// TIA Portal project "000_empty" (V21)

(* hardware
DEVICE "PLC_1"  S7-1500 station
   slot 0: "Rail_0"  Rack  6ES7 590-1***0-0AA0
   slot 1: "PLC_1"  CPU 1513-1 PN  6ES7 513-1AL02-0AB0  V2.9
      slot 3: "CPU display_1"  6ES7591-1AA00-0AA0
      slot 32768: "PROFINET interface_1"  X1
         slot 32769: "Port_1"  X1 P1
         slot 32770: "Port_2"  X1 P2
      slot 34817: "Virtual CP interface port_1"  Virtual CP interface port  Virtual CP interface port
*)

// ===== PLC "PLC_1"  CPU 1513-1 PN =====

VAR_GLOBAL   // PLC tag table "Default tag table"
   "tBool" AT %M0.0 : Bool;
   "tBool2" AT %M0.1 : Bool;
   "tInt" AT %MW2 : Int;
   "tDInt" AT %MD4 : DInt;
   "tReal" AT %MD8 : Real;
   "tWord" AT %MW12 : Word;
   "tByte" AT %MB14 : Byte;
   "tDWord" AT %MD16 : DWord;
   "tTime" AT %MD20 : Time;
   "tIn" AT %I0.0 : Bool;
   "tOut" AT %Q0.0 : Bool;
   "tUInt" AT %MW24 : UInt;
   "tLReal" AT %MD26 : LReal;
   "Tag_1" AT %MW100 : Word;
   "Tag_2" AT %M10.3 : Bool;
   "Tag_3" AT %Q1.0 : Bool;
   "Tag_4" AT %I1.0 : Bool;
   "Tag_5" AT %MD104 : DWord;
   "Tag_6" AT %MB110 : Byte;
   "Tag_7" AT %IW0 : Word;
   "Tag_8" AT %QW0 : Word;
END_VAR

VAR_GLOBAL CONSTANT   // PLC tag table "Default tag table"
   "MAX_COUNT" : Int := 100;
   "GAIN" : Real := 2.5;
   "TXT" : String := 'abc';
END_VAR

TYPE "UDT_Motor"
   STRUCT
      Running : Bool;   // Motor on
      Speed : Real := 1500.0;   // Speed setpoint
      Count : Int := 7;
   END_STRUCT;
END_TYPE

DATA_BLOCK "DB_Global"   // DB1
{ S7_Optimized_Access := 'TRUE' }
   VAR
      xBool : Bool := TRUE;   // Bool comment
      iInt : Int := 42;
      rReal : Real := 3.5;   // Real comment
      aInt : Array[0..3] of Int;
      sData : Struct
         "a" : Bool;
         "b" : DInt := -5;
      END_STRUCT;
   END_VAR
BEGIN
   aInt[1] := 11;
END_DATA_BLOCK

DATA_BLOCK "FB_Empty_DB"   // DB2
{ S7_Optimized_Access := 'TRUE' }
VERSION : 0.1
// stored: InstanceOfName FB_Empty
"FB_Empty"
BEGIN
END_DATA_BLOCK

DATA_BLOCK "DB_Motor"   // DB4
{ S7_Optimized_Access := 'TRUE' }
   VAR
      motor : "UDT_Motor";
   END_VAR
BEGIN
   motor.Speed := 750.0;
END_DATA_BLOCK

DATA_BLOCK "FB_Iface_DB"   // DB5
{ S7_Optimized_Access := 'TRUE' }
VERSION : 0.1
// stored: InstanceOfName FB_Iface
"FB_Iface"
BEGIN
   stInt := 99;
   stBool := TRUE;
END_DATA_BLOCK

DATA_BLOCK "DB_Std"   // DB6
{ S7_Optimized_Access := 'FALSE' }
   VAR
      x : Bool;
      i : Int;
      d : DInt;
      r : Real;
      "by" : Byte;
   END_VAR
BEGIN
END_DATA_BLOCK

// folder: BlockGroup_1

DATA_BLOCK "DB_InGroup"   // DB3
{ S7_Optimized_Access := 'TRUE' }
   VAR
      wWord : Word := 16#00FF;
   END_VAR
BEGIN
END_DATA_BLOCK

// folder: (top level)

DATA_BLOCK "TO_Speed_5_0"   // DB8, Motion_DB
{ S7_Optimized_Access := 'TRUE' }
AUTHOR : SIMATIC
FAMILY : MC_1500
VERSION : 5.0
// stored: InstanceOfName TO_SpeedAxis
"TO_SpeedAxis"
BEGIN
END_DATA_BLOCK

DATA_BLOCK "TO_Posit_6_0"   // DB10, Motion_DB
{ S7_Optimized_Access := 'TRUE' }
AUTHOR : SIMATIC
FAMILY : MC_1500
VERSION : 6.0
// stored: InstanceOfName TO_PositioningAxis
"TO_PositioningAxis"
BEGIN
END_DATA_BLOCK

DATA_BLOCK "TO_Exter_6_0"   // DB13, Motion_DB
{ S7_Optimized_Access := 'TRUE' }
AUTHOR : SIMATIC
FAMILY : MC_1500
VERSION : 6.0
// stored: InstanceOfName TO_ExternalEncoder
"TO_ExternalEncoder"
BEGIN
END_DATA_BLOCK

DATA_BLOCK "SpeedAx_6_0"   // DB14, Motion_DB
{ S7_Optimized_Access := 'TRUE' }
AUTHOR : SIMATIC
FAMILY : MC_1500
VERSION : 6.0
// stored: InstanceOfName TO_SpeedAxis
"TO_SpeedAxis"
BEGIN
END_DATA_BLOCK

FUNCTION_BLOCK "FB_Empty"   // FB1, SCL
{ S7_Optimized_Access := 'TRUE' }
VERSION : 0.1
BEGIN
END_FUNCTION_BLOCK

FUNCTION_BLOCK "FB_Iface"   // FB2, SCL
{ S7_Optimized_Access := 'TRUE' }
VERSION : 0.1
   VAR_INPUT
      iBool : Bool;   // Input bool
      iInt : Int;   // Input int
      iReal : Real;   // Input real
      iArr : Array[0..3] of Int;   // Input array
      iMotor : "UDT_Motor";   // Input UDT
   END_VAR
   VAR_OUTPUT
      oBool : Bool;   // Output bool
      oInt : Int;   // Output int
   END_VAR
   VAR_IN_OUT
      ioReal : Real;   // InOut real
   END_VAR
   VAR
      stInt : Int := 42;   // Static int
      stBool : Bool;   // Static bool comment
   END_VAR
   VAR_TEMP
      tInt : Int;   // Temp int
   END_VAR
   VAR CONSTANT
      cInt : Int := 7;   // Constant int
   END_VAR
BEGIN
   #tInt := #iInt + #cInt;
           #oInt := #tInt;
           #oBool := #iBool;
           #ioReal := #ioReal + #iReal;
END_FUNCTION_BLOCK

FUNCTION_BLOCK "FB_SclCalls"   // FB3, SCL
{ S7_Optimized_Access := 'TRUE' }
VERSION : 0.1
   VAR_INPUT
      start : Bool;
      pt : Time;
   END_VAR
   VAR_OUTPUT
      q : Bool;
      cnt : Int;
   END_VAR
   VAR
      tonInst : TON_TIME;
      tofInst : TOF_TIME;
      tpInst : TP_TIME;
      ctuInst : CTU_INT;
      trig : R_TRIG;
      ftrig : F_TRIG;
      "counter" : Int;
      ifc : "FB_Iface";
   END_VAR
   VAR_TEMP
      r : Real;
      "b" : Bool;
      res : Int;
      tot : Int;
   END_VAR
BEGIN
   #tonInst(IN := #start, PT := #pt);
   #q := #tonInst.Q;
   #tofInst(IN := #start, PT := T#2s);
   #tpInst(IN := #start, PT := #pt, Q => #b);
   #ctuInst(CU := #start, R := FALSE, PV := 10);
   #cnt := #ctuInst.CV;
   #trig(CLK := #start);
   IF #trig.Q THEN
       #counter := 0;
   END_IF;
   #ftrig(CLK := #start);
   #b := #ftrig.Q;
   #ifc(iBool := TRUE, iInt := 2, iReal := 1.0, ioReal := #r);
   #cnt := #ifc.oInt;
   "FB_Iface_DB"(iBool := #start, iInt := #cnt, iReal := #r, ioReal := #r, oInt => #cnt);
   "FC_SclOps"();
   #res := "FC_SclCtl"(n := 5, flag := TRUE, total => #tot);
   #res := "FC_SclCtl"(n := #res, flag := #b, total => #tot);
END_FUNCTION_BLOCK

FUNCTION_BLOCK "FB_SclLocal"   // FB4, SCL
{ S7_Optimized_Access := 'TRUE' }
VERSION : 0.1
   VAR_INPUT
      start : Bool;
   END_VAR
   VAR_IN_OUT
      io : Int;
   END_VAR
   VAR
      "counter" : Int;
      arr : Array[0..9] of Int;
      arr2 : Array[1..3, 1..4] of Real;
      mot : "UDT_Motor";
      st : Struct
         "a" : Int;
         "b" : Real;
         c : Array[0..2] of Bool;
      END_STRUCT;
   END_VAR
   VAR_TEMP
      i : Int;
   END_VAR
BEGIN
   #arr[0] := 1;
   #arr[#i] := #arr[#i + 1] + #io;
   #arr2[2, 3] := 1.5;
   #st.a := 10;
   #st.b := #st.a;
   #st.c[1] := TRUE;
   #mot.Speed := 100.0;
   #mot.Running := #st.c[0];
   #counter += 1;
   #io := #counter;
END_FUNCTION_BLOCK

FUNCTION_BLOCK "FB_LadTech"   // FB5, LAD
{ S7_Optimized_Access := 'TRUE' }
   VAR_INPUT
      sp : Real;
      pv : Real;
   END_VAR
   VAR_OUTPUT
      outv : Real;
      err : Bool;
   END_VAR
BEGIN

REGION Network 1: PID call
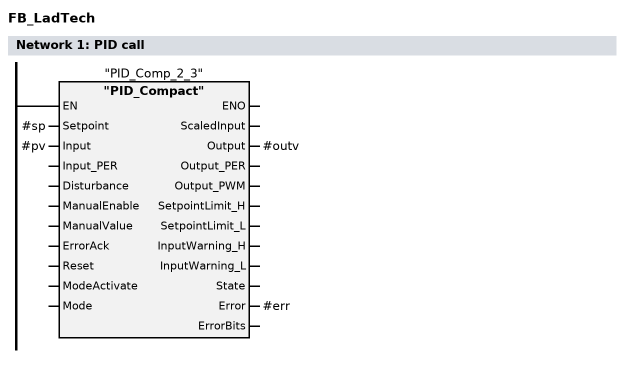
   RUNG wire#powerrail
      "PID_Comp_2_3"(Setpoint := #sp, Input := #pv, Output => #outv, Error => #err, Input_PER :=, Disturbance :=, ManualEnable :=, ManualValue :=, ErrorAck :=, Reset :=, ModeActivate :=, ScaledInput =>, Output_PER =>, Output_PWM =>, SetpointLimit_H =>, SetpointLimit_L =>, InputWarning_H =>, InputWarning_L =>, State =>, ErrorBits =>, Mode :=)
   END_RUNG
   // the same network as SCL:
   "PID_Comp_2_3"(Setpoint := #sp, Input := #pv, Output => #outv, Error => #err);   // "PID_Compact"
END_REGION
END_FUNCTION_BLOCK

FUNCTION_BLOCK "FB_FbdTech"   // FB6, FBD
{ S7_Optimized_Access := 'TRUE' }
   VAR_INPUT
      sp : Real;
      pv : Real;
   END_VAR
   VAR_OUTPUT
      outv : Real;
      err : Bool;
   END_VAR
BEGIN

REGION Network 1: PID call
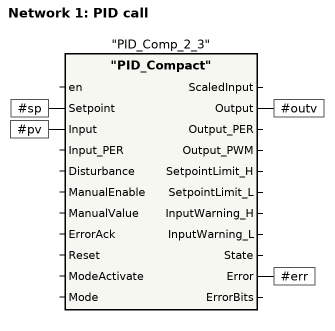
   "PID_Comp_2_3"(Setpoint := #sp, Input := #pv, Output => #outv, Error => #err);   // "PID_Compact"
END_REGION
END_FUNCTION_BLOCK

FUNCTION_BLOCK "FB_SclTech"   // FB7, SCL
{ S7_Optimized_Access := 'TRUE' }
   VAR_INPUT
      sp : Real;
      pv : Real;
   END_VAR
   VAR_OUTPUT
      outv : Real;
      err : Bool;
   END_VAR
BEGIN
// PID call
   "PID_Comp_2_3"(Setpoint := #sp, Input := #pv, Output => #outv, Error => #err);
END_FUNCTION_BLOCK

FUNCTION "FC_SclOps" : Void   // FC1, SCL
{ S7_Optimized_Access := 'TRUE' }
VERSION : 0.1
   VAR_TEMP
      b1 : Bool;
      b2 : Bool;
      b3 : Bool;
      i1 : Int;
      i2 : Int;
      i3 : Int;
      d1 : DInt;
      r1 : Real;
      r2 : Real;
      l1 : LReal;
      w1 : Word;
      w2 : Word;
      dw1 : DWord;
      by1 : Byte;
      u1 : UInt;
   END_VAR
BEGIN
   // arithmetic
           #i1 := 1 + 2 - 3 * 4;
           #i2 := #i1 / 2;
           #i3 := #i1 MOD 3;
           #r1 := #r2 ** 2.0;
           #i1 := -#i2;
           #i1 := +#i2;
           #i1 := (#i2 + #i3) * (#i2 - #i3);
           #d1 := #i1 * #i2;
           #r1 := #r2 / 3.0;
           #u1 := 5;
           // logic
           #b1 := NOT #b2;
           #b1 := #b2 AND #b3;
           #b1 := #b2 OR #b3;
           #b1 := #b2 XOR #b3;
           #b1 := #b2 & #b3;
           #b1 := (#b2 AND #b3) OR NOT (#b2 XOR #b3);
           #w1 := #w1 AND #w2;
           #w1 := #w1 OR #w2;
           #w1 := #w1 XOR #w2;
           #w1 := NOT #w2;
           // comparison
           #b1 := #i1 = #i2;
           #b1 := #i1 <> #i2;
           #b1 := #i1 < #i2;
           #b1 := #i1 <= #i2;
           #b1 := #i1 > #i2;
           #b1 := #i1 >= #i2;
           #b1 := #r1 > 1.5 AND #r2 <= 2.5;
           // compound assignment
           #i1 += 1;
           #i1 -= 1;
           #i1 *= 2;
           #i1 /= 2;
           // mixed types
           #l1 := #r1 + #d1;
           #r1 := #i1;
           #by1 := 16#FF;
           #dw1 := 16#DEADBEEF;
           #w1 := 2#1010_1010;
           #i1 := 8#17;
           #r1 := 1.0E3;
           #r2 := 2.5e-3;
           #l1 := 3.141592653589793;
END_FUNCTION

FUNCTION "FC_SclCtl" : Int   // FC2, SCL
{ S7_Optimized_Access := 'TRUE' }
VERSION : 0.1
   VAR_INPUT
      n : Int;
      flag : Bool;
   END_VAR
   VAR_OUTPUT
      total : Int;
   END_VAR
   VAR_TEMP
      i : Int;
      j : Int;
      x : Int;
      "b" : Bool;
   END_VAR
BEGIN
   (* block comment
      over two lines *)
   #total := 0;
   // IF forms
   IF #flag THEN
       #total := 1;
   END_IF;
   IF #n > 5 THEN
       #total := 2;
   ELSE
       #total := 3;
   END_IF;
   IF #n > 10 THEN
       #total := 4;
   ELSIF #n > 5 THEN
       #total := 5;
   ELSIF #n > 0 THEN
       #total := 6;
   ELSE
       #total := 7;
   END_IF;
   // CASE
   CASE #n OF
       0:
           #total := 10;
       1, 2:
           #total := 11;
       3..5:
           #total := 12;
       6, 8..9:
           #total := 13;
   ELSE
       #total := 14;
   END_CASE;
   CASE #x OF
       1:
           ;
   END_CASE;
   // FOR with BY, EXIT, CONTINUE
   FOR #i := 0 TO 10 DO
       #total += #i;
   END_FOR;
   FOR #i := 10 TO 0 BY -2 DO
       IF #i = 4 THEN
           CONTINUE;
       END_IF;
       IF #i = 2 THEN
           EXIT;
       END_IF;
       #total += #i;
   END_FOR;
   // nested loops
   FOR #i := 1 TO 3 DO
       FOR #j := 1 TO 3 DO
           #total := #total + #i * #j;
       END_FOR;
   END_FOR;
   // WHILE
   #x := 0;
   WHILE #x < 5 DO
       #x := #x + 1;
   END_WHILE;
   // REPEAT
   REPEAT
       #x := #x - 1;
   UNTIL #x <= 0
   END_REPEAT;
   // REGION
   REGION Calculation
       #total := #total * 2;
   END_REGION;
   // GOTO and labels
   IF #flag THEN
       GOTO done;
   END_IF;
   #total := #total + 1;
   done:
   #b := TRUE;
   // empty statement and RETURN
   ;
   #FC_SclCtl := #total;
   RETURN;
END_FUNCTION

FUNCTION "FC_SclLit" : Void   // FC3, SCL
{ S7_Optimized_Access := 'TRUE' }
VERSION : 0.1
   VAR_TEMP
      "b" : Bool;
      "by" : Byte;
      w : Word;
      dw : DWord;
      lw : LWord;
      si : SInt;
      i : Int;
      di : DInt;
      li : LInt;
      usi : USInt;
      ui : UInt;
      udi : UDInt;
      uli : ULInt;
      r : Real;
      lr : LReal;
      t : Time;
      lt : LTime;
      d : Date;
      tod : Time_Of_Day;
      ltod : LTime_Of_Day;
      "dt" : DTL;
      ldt : LDT;
      c : Char;
      wc : WChar;
      s : String;
      ws : WString;
      sn : String[10];
   END_VAR
BEGIN
   #b := TRUE;
           #b := FALSE;
           #by := 16#7F;
           #w := 16#BEEF;
           #dw := 16#DEAD_BEEF;
           #lw := 16#0123_4567_89AB_CDEF;
           #si := -128;
           #i := 32767;
           #di := -2147483648;
           #li := 9223372036854775807;
           #usi := 255;
           #ui := 65535;
           #udi := 4294967295;
           #uli := 18446744073709551615;
           #r := 3.5;
           #r := 1.0e10;
           #lr := 2.718281828459045;
           #t := T#5s;
           #t := T#1d_2h_3m_4s_5ms;
           #t := T#-10s;
           #lt := LT#1d2h3m4s5ms6us7ns;
           #d := D#2024-02-29;
           #tod := TOD#12:30:45.123;
           #ltod := LTOD#23:59:59.999999999;
           #dt := DTL#2024-02-29-12:30:45.5;
           #ldt := LDT#2024-02-29-12:30:45;
           #c := 'A';
           #c := '$N';
           #wc := WCHAR#'W';
           #s := 'Hello';
           #s := 'It$'s a $$ test';
           #s := '';
           #ws := WSTRING#'Wide';
           #sn := 'abc';
           #i := INT#5;
           #di := DINT#-5;
           #r := REAL#2.5;
           #w := WORD#16#FF;
           #by := BYTE#16#0F;
           #b := BOOL#1;
           #t := TIME#10s;
           #lr := LREAL#1.0;
           #i := 1_000;
END_FUNCTION

FUNCTION "FC_SclGlobal" : Void   // FC4, SCL
{ S7_Optimized_Access := 'TRUE' }
VERSION : 0.1
   VAR_TEMP
      i : Int;
   END_VAR
BEGIN
   "DB_Global".iInt := 5;
   "DB_Global".xBool := NOT "DB_Global".xBool;
   "DB_Global".aInt[2] := "DB_Global".aInt[1] + 1;
   "DB_Global".aInt[#i] := 0;
   "DB_Global".sData.b := "DB_Global".sData.b + 1;
   "DB_Motor".motor.Speed := "DB_Motor".motor.Speed * 2.0;
   "FB_Iface_DB".stInt := 3;
   "FB_Iface_DB".iArr[1] := 4;
   "FB_Iface_DB".iMotor.Speed := 5.0;
   "tInt" := "tInt" + 1;
   "tBool" := "tIn" AND NOT "tBool2";
   "tOut" := "tBool";
   "tReal" := "tReal" * 0.5;
END_FUNCTION

FUNCTION "FC_SclAbs" : Void   // FC5, SCL
{ S7_Optimized_Access := 'TRUE' }
VERSION : 0.1
   VAR_TEMP
      "b" : Bool;
   END_VAR
BEGIN
   "Tag_1" := 5;
   "Tag_2" := TRUE;
   "Tag_3" := "Tag_4";
   "Tag_5" := 100;
   "Tag_6" := 1;
   #b := "Tag_2";
END_FUNCTION

FUNCTION "FC_SclSlice" : Void   // FC6, SCL
{ S7_Optimized_Access := 'TRUE' }
VERSION : 0.1
   VAR_TEMP
      "b" : Bool;
      w : Word;
      dw : DWord;
      "by" : Byte;
      lw : LWord;
      i : Int;
   END_VAR
BEGIN
   #b := #w.%X3;
   #w.%X0 := TRUE;
   #by := #w.%B1;
   #w.%B0 := #by;
   #dw.%W1 := #w;
   #b := #dw.%X31;
   #w := #dw.%W0;
   #by := #dw.%B3;
   #dw.%B2 := #by;
   #b := #lw.%X63;
   #w := #lw.%W3;
   #dw := #lw.%D1;
   "tWord".%X5 := #b;
   #b := "tDWord".%X7;
END_FUNCTION

FUNCTION "FC_SclMath" : Void   // FC7, SCL
{ S7_Optimized_Access := 'TRUE' }
VERSION : 0.1
   VAR_TEMP
      i : Int;
      j : Int;
      d : DInt;
      r : Real;
      r2 : Real;
      lr : LReal;
      "b" : Bool;
      w : Word;
      dw : DWord;
      "by" : Byte;
      t : Time;
   END_VAR
BEGIN
   #r := ABS(#r2);
   #r := SQRT(#r2);
   #r := SQR(#r2);
   #r := LN(#r2);
   #r := EXP(#r2);
   #r := SIN(#r2);
   #r := COS(#r2);
   #r := TAN(#r2);
   #r := ASIN(#r2);
   #r := ACOS(#r2);
   #r := ATAN(#r2);
   #i := ABS(#j);
   #i := MIN(IN1 := #i, IN2 := #j);
   #i := MAX(IN1 := #i, IN2 := #j);
   #i := LIMIT(MN := 0, IN := #i, MX := 100);
   #i := MIN(IN1 := #i, IN2 := #j, IN3 := 5);
   #i := MAX(IN1 := #i, IN2 := #j, IN3 := 5);
   #i := SEL(G := #b, IN0 := #i, IN1 := #j);
   #i := MUX(K := #j, IN0 := 1, IN1 := 2, IN2 := 3);
   #r := INT_TO_REAL(#i);
   #i := REAL_TO_INT(#r);
   #d := REAL_TO_DINT(#r);
   #i := DINT_TO_INT(#d);
   #d := INT_TO_DINT(#i);
   #d := TRUNC(#r);
   #d := ROUND(#r);
   #d := CEIL(#r);
   #d := FLOOR(#r);
   #r := DINT_TO_REAL(#d);
   #w := INT_TO_WORD(#i);
   #i := WORD_TO_INT(#w);
   #dw := SHL(IN := #dw, N := 2);
   #dw := SHR(IN := #dw, N := 2);
   #dw := ROL(IN := #dw, N := 1);
   #dw := ROR(IN := #dw, N := 1);
   #w := SHL(IN := #w, N := 1);
   #by := BYTE#16#01;
   #t := INT_TO_TIME(#i);
   #r := NORM_X(MIN := 0, VALUE := #i, MAX := 27648);
   #i := SCALE_X(MIN := 0, VALUE := #r, MAX := 27648);
   #d := DWORD_TO_DINT(#dw);
   #dw := DINT_TO_DWORD(#d);
   #r := FRAC(#r2);
END_FUNCTION

FUNCTION "FC_SclStr" : Void   // FC8, SCL
{ S7_Optimized_Access := 'TRUE' }
VERSION : 0.1
   VAR_TEMP
      s : String;
      s2 : String;
      ws : WString;
      i : Int;
      c : Char;
      "b" : Bool;
      r : Real;
   END_VAR
BEGIN
   #i := LEN(#s);
   #s := CONCAT(IN1 := #s, IN2 := #s2);
   #s := LEFT(IN := #s, L := 2);
   #s := RIGHT(IN := #s, L := 2);
   #s := MID(IN := #s, L := 2, P := 1);
   #i := FIND(IN1 := #s, IN2 := #s2);
   #s := INSERT(IN1 := #s, IN2 := #s2, P := 1);
   #s := DELETE(IN := #s, L := 1, P := 1);
   #s := REPLACE(IN1 := #s, IN2 := #s2, L := 1, P := 1);
   #b := #s = #s2;
   #b := #s <> #s2;
   #b := #s < #s2;
   #c := #s[1];
   #s[1] := #c;
   #s := INT_TO_STRING(#i);
   #i := STRING_TO_INT(#s);
   #s := REAL_TO_STRING(#r);
   #ws := STRING_TO_WSTRING(#s);
END_FUNCTION

FUNCTION "FC_SclMisc" : Void   // FC9, SCL
{ S7_Optimized_Access := 'TRUE' }
VERSION : 0.1
   VAR_IN_OUT
      arr : Array[1..2, 1..2] of Int;
      arr3 : Array[0..1, 0..1, 0..1] of Int;
   END_VAR
   VAR_TEMP
      i : Int;
      d : DInt;
      "b" : Bool;
      v : Variant;
      "by" : Byte;
      w : Word;
      p : Int;
   END_VAR
BEGIN
   #by := PEEK(area := 16#84, dbNumber := 1, byteOffset := 0);
   POKE(area := 16#84, dbNumber := 1, byteOffset := 0, value := #by);
   #w := PEEK_WORD(area := 16#84, dbNumber := 1, byteOffset := 0);
   POKE(area := 16#84, dbNumber := 1, byteOffset := 0, value := #w);
   #b := PEEK_BOOL(area := 16#84, dbNumber := 1, byteOffset := 0, bitOffset := 1);
   #v := REF("DB_Global".iInt);
   #arr[1, 1] := 1;
   #arr3[0, 1, 0] := 3;
   #b := IS_ARRAY(#v);
   #i := CountOfElements(#v);
   #d := #i;
END_FUNCTION

FUNCTION "FC_SclArr" : Void   // FC10, SCL
{ S7_Optimized_Access := 'TRUE' }
VERSION : 0.1
   VAR_IN_OUT
      arr : Array[1..2, 1..2] of Int;
      arr3 : Array[0..1, 0..1, 0..1] of Int;
   END_VAR
   VAR_TEMP
      i : Int;
   END_VAR
BEGIN
   #arr[#i, 1] := #arr[1, #i];
   #arr3[#i, 0, 1] := #arr3[1, #i, 0];
END_FUNCTION

FUNCTION "FC_SclAbs2" : Void   // FC11, SCL
{ S7_Optimized_Access := 'TRUE' }
VERSION : 0.1
   VAR_TEMP
      "b" : Bool;
      i : Int;
      d : DInt;
      r : Real;
   END_VAR
BEGIN
   %DB6.DBX0.0 := TRUE;
           #b := %DB6.DBX0.0;
           %DB6.DBW2 := 5;
           #i := %DB6.DBW2;
           %DB6.DBD4 := 7;
           #d := %DB6.DBD4;
           %DB6.DBB8 := 3;
           "DB_Std".x := #b;
           "DB_Std".i := #i;
           "DB_Std".r := #r;
           #i := "DB_Std".i + 1;
END_FUNCTION

FUNCTION "FC_SclVar" : Void   // FC12, SCL
{ S7_Optimized_Access := 'TRUE' }
VERSION : 0.1
   VAR_INPUT
      v : Variant;
   END_VAR
   VAR_TEMP
      i : Int;
      "b" : Bool;
      n : UDInt;
      t : Time;
      w : Word;
   END_VAR
BEGIN
   #n := CountOfElements(#v);
           #b := IS_ARRAY(#v);
           #b := TypeOf(#v) = TypeOf(#i);
           VariantGet(SRC := #v, DST => #i);
           VariantPut(SRC := #i, DST := #v);
           #i := MOVE_BLK_VARIANT(SRC := #v, COUNT := 1, SRC_INDEX := 0, DEST_INDEX := 0, DEST => #v);
           #b := ENO;

       #i := 1;    // tab-separated

           #i := 2;
END_FUNCTION

FUNCTION "FC_SclMore" : Void   // FC13, SCL
{ S7_Optimized_Access := 'TRUE' }
VERSION : 0.1
   VAR_INPUT
      "my var" : Int;
   END_VAR
   VAR_IN_OUT
      va : Array[*] of Int;
   END_VAR
   VAR_TEMP
      i : Int;
      j : Int;
      d : DInt;
      t1 : Time;
      t2 : Time;
      dt1 : Date;
      dt2 : Date;
      tod : Time_Of_Day;
      r : Real;
      s : String;
      ws : WString;
      "b" : Bool;
      w : Word;
      tcnt : DInt;
   END_VAR
   VAR CONSTANT
      cMax : Int := 10;
      cText : String := 'const';
   END_VAR
BEGIN
   // quoted identifiers, user constants
   #i := #"my var" + "MAX_COUNT";
   #r := "GAIN" * 2.0;
   #s := "TXT";
   #i := #cMax;
   #s := #cText;
   // several statements per line
   #i := 1; #j := 2; #d := 3;
   // trailing and inline comments
   #i := 1; // trailing comment
   #j := 1 (* inline *) + 2;
   (* single line block comment *)
   (* a *) #i := 3; (* b *)
   // time and date arithmetic
   #t1 := #t1 + #t2;
   #t1 := #t1 - T#1s;
   #t1 := #t1 * 2;
   #t1 := #t1 / 2;
   #tod := #tod + #t1;
   #b := #t1 > #t2;
   #b := #dt1 <= #dt2;
   #tcnt := UPPER_BOUND(ARR := #va, DIM := 1);
   #tcnt := LOWER_BOUND(ARR := #va, DIM := 1);
   // arrays of UDT and nested access
   "DB_Motor".motor.Speed := 1.0;
   "FB_Iface_DB".iArr[#i] := #j;
   // peripheral and direct I/O
   #w := "Tag_7":P;
   "Tag_8":P := #w;
   #b := "tIn";
   // unicode
   #s := 'äöü ß € ünï';
   #ws := WSTRING#'äöü €';
   // long expression
   #r := (((#r + 1.0) * (#r - 1.0)) / ((#r + 2.0) * (#r - 2.0))) + (((#r + 3.0) * (#r - 3.0)) / ((#r + 4.0) * (#r - 4.0)));
   // nested structured statements
   IF #b THEN
       FOR #i := 0 TO 3 DO
           WHILE #j < 10 DO
               CASE #j OF
                   1:
                       #j += 1;
                   2..4:
                       REPEAT
                           #j += 2;
                       UNTIL #j > 5
                       END_REPEAT;
               ELSE
                   #j += 3;
               END_CASE;
           END_WHILE;
       END_FOR;
   ELSIF NOT #b THEN
       REGION Outer
           REGION Inner
               #i := 0;
           END_REGION;
       END_REGION;
   END_IF;
   FOR #i := #j TO #d BY #i DO
       #j := #i;
   END_FOR;
END_FUNCTION

ORGANIZATION_BLOCK "Main"   // OB1, LAD, ProgramCycle
TITLE = "Main Program Sweep (Cycle)"
{ S7_Optimized_Access := 'TRUE' }
VERSION : 0.1
   VAR_INPUT
      Initial_Call : Bool;   // Initial call of this OB
      Remanence : Bool;   // =True, if remanent data are available
   END_VAR
BEGIN
END_ORGANIZATION_BLOCK